Staubli VAL3: getSize.pgx

public program getSize(num& x_nSize)
begin
   if size(progTemp:pProgItem)>0
    x_nSize=size(progTemp:pProgItem)
  else
    x_nSize=1
  endIf
end
